(* IEC 61131-3 sources: Cocktail-Mix-Maschine-V2/Code für SPS/Logical/Library, 1 file *)

(* ---- Library.fun ---- *)
{REDUND_ERROR} FUNCTION setOutputs : BOOL (*TODO: Add your comment here*) (*$GROUP=User,$CAT=User,$GROUPICON=User.png,$CATICON=User.png*)
	VAR_INPUT
		ventil1 : BOOL;
		ventil2 : BOOL;
		ventil3 : BOOL;
		ventil4 : BOOL;
		ventil5 : BOOL;
		ventil6 : BOOL;
		ventil7 : BOOL;
		ventil8 : BOOL;
		rot : BOOL;
		gruen : BOOL;
		pumpe : BOOL;
		motor : BOOL;
	END_VAR
END_FUNCTION
